// TIA Portal V19 export
DATA_BLOCK "CONTROL_DB"   // DB9
// stored: InstanceOfName SEMI/_AUTO, InstanceOfType FB
"SEMI/_AUTO"
   // VAR_INPUT
   //    SEMI_AUTO : Bool;
   //    UCHWS_IN : Bool;
   //    CHWS_IN : Bool;
   //    CTS_IN : Bool;
   //    HWS_IN : Bool;
   //    HMI_SEMI_SEL : Int;
   // END_VAR
   // VAR_OUTPUT
   //    UCHW_CMD : Bool;
   //    CHW_CMD : Bool;
   //    CT_CMD : Bool;
   //    HW_CMD : Bool;
   // END_VAR
   // VAR
   //    "STEP" : Int;
   // END_VAR
BEGIN
END_DATA_BLOCK
